// TIA Portal V20 export
// export: Created 2025-07-07T08:55:10.1278921Z, ExportSetting None, DisplayName Totally Integrated Automation Portal, DisplayVersion V20 Update 5, DisplayName TIA Portal Openness, DisplayVersion V20 Update 5, DisplayName TIA Portal Version Control Interface, DisplayVersion V20, DisplayName SINAMICS Startdrive Advanced, DisplayVersion V20, DisplayName SINAMICS Startdrive G130, G150, S120, S150, SINAMICS MV, S210, DisplayVersion V20, DisplayName SINAMICS Startdrive G110M, G120, G120C, G120D, G120P, G115D, DisplayVersion V20, DisplayName STEP 7 Professional, DisplayVersion V20 Update 5, DisplayName STEP 7 Safety, DisplayVersion V20, DisplayName WinCC Advanced, DisplayVersion V20 Update 5
DATA_BLOCK "FB_PR_GantryUnload_Seqv25_DB"   // DB1
// stored: InstanceOfName FB_PR_GantryUnload_Seqv25, InstanceOfType FB
"FB_PR_GantryUnload_Seqv25"
   // VAR_INPUT
   //    iAutoRunning : Bool;
   //    iCenteringSlideAtHome : Bool;
   //    iCenteringSlideAtWork : Bool;
   //    iDistSenHighLimit : Int;
   //    iDistSenLowLimit : Int;
   //    iDistSensorIP : Int;
   //    iDryCycleWithoutPal : Bool;
   //    iGantryOutofZone : Bool;
   //    iGantryPickOver : Bool;
   //    iPCAckZero : Bool;
   //    iPCBypass : Bool;
   //    iPCDataReadOver : Bool;
   //    iPCDataWriteOver : Bool;
   //    iPalletPresent : Bool;
   //    iProcessStart : Bool;
   //    iReset_fault : Bool;
   //    iRetryPB : Bool;
   //    iScanErr : Bool;
   //    iScanOver : Bool;
   //    iScannerBypass : Bool;
   //    iSstMode : Bool;
   //    iSstPB : Bool;
   // END_VAR
   // VAR_OUTPUT
   //    qCenteringSlideAdvance : Bool;
   //    qCenteringSlideRetract : Bool;
   //    qCheckDistance : Bool;
   //    qGantryOkToUnload : Bool;
   //    qMsg : Array[0..2] of Bool;
   //    qPCReadCmd : Bool;
   //    qPCUploadCmd : Bool;
   //    qProcessOver : Bool;
   //    qScanCmd : Bool;
   // END_VAR
BEGIN
END_DATA_BLOCK
